TYPE ET_CalcExtTiltState :
(
	ET_CalcExtTiltState_eWaitExecute := 0,
	ET_CalcExtTiltState_eCalcTiltPos := 5,
	ET_CalcExtTiltState_eDone := 197,
	ET_CalcExtTiltState_eError := 198,
	ET_CalcExtTiltState_eNoExecute := 199
);
END_TYPE

(* stored: Version 1.1.0.1, ProductVersion 3.1.4024.15
   DUT ET_CalcExtTiltState: Id {3b384982-2175-4d3f-8c54-37296742cebc} *)
